FUNCTION_BLOCK FB_IoGroup IMPLEMENTS I_IoGroup

VAR
	aIoArray	: ARRAY [1..30] OF I_IoBase;
	nIoIndex	: INT := 0;
END_VAR

Update();


METHOD AddIo
VAR_INPUT
	bIo	: I_IoBit;
END_VAR
IF bIo <> 0 THEN
	nIoIndex  := nIoIndex + 1;
	aIoArray[nIoIndex] := bIo;
	
END_IF
END_METHOD


METHOD Update
VAR
    i : INT;
END_VAR
FOR i := 1 TO nIoIndex DO
	aIoArray[i].Update();
	
END_FOR
END_METHOD

END_FUNCTION_BLOCK

(* stored: Version 1.1.0.1
   POU FB_IoGroup: Id {384c065e-b6a2-4bce-804b-2301a51c0a14}, SpecialFunc None
   Method AddIo: Id {f63768c2-3bfe-411c-aabc-594490ffa8e1}
   Method Update: Id {d71c24d0-f573-417c-b717-61ca25a7712e} *)
